FUNCTION F_EL6910MessageTemplate : STRING(255)
VAR_INPUT
    wTextId : WORD;
END_VAR

CASE wTextId OF
    16#0001: F_EL6910MessageTemplate := 'Primary MC: GLOBAL_Fault with Code 0x%x and Additional Code 0x%x';
    16#0002: F_EL6910MessageTemplate := 'Primary MC: GLOBAL_Shutdown with Code 0x%x and Additional Code 0x%x';
    16#0003: F_EL6910MessageTemplate := 'Secondary MC: GLOBAL_Fault with Code 0x%x and Additional Code 0x%x';
    16#0004: F_EL6910MessageTemplate := 'Secondary MC: GLOBAL_Shutdown with Code 0x%x and Additional Code 0x%x';
    16#0005: F_EL6910MessageTemplate := 'Primary MC: Stored GLOBAL_Fault with Code 0x%x and Additional Code 0x%x';
    16#0006: F_EL6910MessageTemplate := 'Secondary MC: Stored GLOBAL_Fault with Code 0x%x and Additional Code 0x%x';
    16#0007: F_EL6910MessageTemplate := 'Diag-Message-Overflow: %d messages got lost';
    16#0008: F_EL6910MessageTemplate := 'Primary MC: the CRC of the FRAM Data was wrong (Diag-Code=%d)';
    16#0009: F_EL6910MessageTemplate := 'Secondary MC: the CRC of the FRAM Data was wrong (Diag-Code=%d)';
    16#0010: F_EL6910MessageTemplate := 'Reserved CfgData has to be zero st offset %d';
    16#0011: F_EL6910MessageTemplate := 'The password is wrong';
    16#0012: F_EL6910MessageTemplate := 'The user was not found';
    16#0013: F_EL6910MessageTemplate := 'The CRC of the login data does not match';
    16#0014: F_EL6910MessageTemplate := 'The serial number of the login data does not match';
    16#0015: F_EL6910MessageTemplate := 'The login watchdog has been expired';
    16#0016: F_EL6910MessageTemplate := 'The user was logged out before';
    16#0017: F_EL6910MessageTemplate := 'The user has not sufficient access rights';
    16#0018: F_EL6910MessageTemplate := 'The reserved area of the CfgData was not 0';
    16#0019: F_EL6910MessageTemplate := 'The CRC of the CfgData was wrong';
    16#001A: F_EL6910MessageTemplate := 'The user name is wrong at word offset 0x%x when changing the password';
    16#001B: F_EL6910MessageTemplate := 'The requested number of users is too big';
    16#001D: F_EL6910MessageTemplate := 'The user update flags are wrong at word offset 0x%x when changing the password';
    16#001E: F_EL6910MessageTemplate := 'The wrong user (user %d) is logged in when changing the password (user %d found in the received data)';
    16#0021: F_EL6910MessageTemplate := 'the maximum Global-Shutdown counter was exceeded in the Vendor Data (maximum value: %d, actual value: %d)';
    16#0030: F_EL6910MessageTemplate := 'Sync Manager 2 Address (0x%x) is invalid, minimum value = 0x%x, maximum value = 0x%x';
    16#0031: F_EL6910MessageTemplate := 'Sync Manager 3 Address (0x%x) is invalid, minimum value = 0x%x, maximum value = 0x%x';
    16#0032: F_EL6910MessageTemplate := 'Sync Manager 4 Address (0x%x) is invalid, minimum value = 0x%x, maximum value = 0x%x';
    16#0033: F_EL6910MessageTemplate := 'Sync Manager 5 Address (0x%x) is invalid, minimum value = 0x%x, maximum value = 0x%x';
    16#0034: F_EL6910MessageTemplate := 'Sync Manager 2 Size (%d) is invalid, minimum value = %d, maximum value = %d';
    16#0035: F_EL6910MessageTemplate := 'Sync Manager 3 Size (%d) is invalid, minimum value = %d, maximum value = %d';
    16#0036: F_EL6910MessageTemplate := 'Sync Manager 4 Size (%d) is invalid, minimum value = %d, maximum value = %d';
    16#0037: F_EL6910MessageTemplate := 'Sync Manager 5 Size (%d) is invalid, minimum value = %d, maximum value = %d';
    16#0038: F_EL6910MessageTemplate := 'Sync Manager %d Settings (Offset 4-7) are invalid, expected values = 0x%x, 0x%x';
    16#0044: F_EL6910MessageTemplate := 'Sync Manager 6 Address (0x%x) is invalid, minimum value = 0x%x, maximum value = 0x%x';
    16#0045: F_EL6910MessageTemplate := 'Sync Manager 7 Address (0x%x) is invalid, minimum value = 0x%x, maximum value = 0x%x';
    16#0048: F_EL6910MessageTemplate := 'Sync Manager 6 Size (%d) is invalid, minimum value = %d, maximum value = %d';
    16#0049: F_EL6910MessageTemplate := 'Sync Manager 7 Size (%d) is invalid, minimum value = %d, maximum value = %d';
    16#0101: F_EL6910MessageTemplate := 'Primary MC: Completed RAM TEST: Starttime: 0x%x and Stoptime: 0x%x . The calculated timediff is 0x%x.';
    16#0102: F_EL6910MessageTemplate := 'Secondary MC: Completed RAM TEST: Starttime: 0x%x and Stoptime: 0x%x . The calculated timediff is 0x%x.';
    16#0115: F_EL6910MessageTemplate := 'Controller %d: Maximum temperature exceeded. Temperature is 0x%x, should be <= 0x%x.';
    16#0116: F_EL6910MessageTemplate := 'Controller %d: Minimum temperature alert. Temperature is 0x%x, should be >= 0x%x.';
    16#0117: F_EL6910MessageTemplate := 'Controller %d: Temperature difference too high. Difference is %d, should be <= %d.';
    16#0118: F_EL6910MessageTemplate := 'Controller %d: Maximum voltage alert (Partner_VCC). Voltage is 0x%x, should be <= 0x%x.';
    16#0119: F_EL6910MessageTemplate := 'Controller %d: Minimum voltage alert (Partner_VCC). Voltage is 0x%x, should be >= 0x%x.';
    16#011A: F_EL6910MessageTemplate := 'Controller %d: Maximum voltage alert (ECAT_VCC). Voltage is 0x%x, should be <= 0x%x.';
    16#011B: F_EL6910MessageTemplate := 'Controller %d: Minimum voltage alert (ECAT_VCC). Voltage is 0x%x, should be >= 0x%x.';
    16#011E: F_EL6910MessageTemplate := 'Controller %d: Timer Tick Difference is too high. Difference is 0x%x, should be >= 0x%x.';
    16#011F: F_EL6910MessageTemplate := 'Controller %d: Minimum value alert (Individual ADC Check). Channel parameter = %d. Actual value is 0x%x.';
    16#0120: F_EL6910MessageTemplate := 'Controller %d: Maximum value alert (Individual ADC Check). Channel parameter = %d. Actual value is 0x%x.';
    16#2001: F_EL6910MessageTemplate := 'The %d. connection has received an invalid FSoE-Cmd in state CONNECTION';
    16#2002: F_EL6910MessageTemplate := 'The %d. connection has received an unknown FSoE-Cmd in state CONNECTION';
    16#2003: F_EL6910MessageTemplate := 'The %d. connection has received an invalid FSoE-ConnID in state CONNECTION';
    16#2004: F_EL6910MessageTemplate := 'The %d. connection has received an invalid FSoE-CRC in state CONNECTION';
    16#2005: F_EL6910MessageTemplate := 'The FSoE-Watchdog of the %d. connection has been expired in state CONNECTION';
    16#2006: F_EL6910MessageTemplate := 'On the %d. connection the received FSoE-Address (0x%x) does not match with the expected FSoE-Address (0x%x)';
    16#2007: F_EL6910MessageTemplate := 'On the %d. connection the received connection data do not match with the sent values';
    16#200C: F_EL6910MessageTemplate := 'On the %d. connection in state CONNECTION the Connection was restarted from the FSoE-Master';
    16#200E: F_EL6910MessageTemplate := 'A Module fault was detected on the %d. connection in state CONNECTION';
    16#2011: F_EL6910MessageTemplate := 'On the %d. connection in state CONNECTION a FSoE-Reset with Error-Code 1 was received which means that the communication partner has received an invalid FSoE-Cmd';
    16#2012: F_EL6910MessageTemplate := 'On the %d. connection in state CONNECTION a FSoE-Reset with Error-Code 2 was received which means that the communication partner has received an unknown FSoE-Cmd';
    16#2013: F_EL6910MessageTemplate := 'On the %d. connection in state CONNECTION a FSoE-Reset with Error-Code 3 was received which means that the communication partner has received an invalid FSoE-ConnID';
    16#2014: F_EL6910MessageTemplate := 'On the %d. connection in state CONNECTION a FSoE-Reset with Error-Code 4 was received which means that the communication partner has received an invalid FSoE-CRC';
    16#2015: F_EL6910MessageTemplate := 'On the %d. connection in state CONNECTION a FSoE-Reset with Error-Code 5 was received which means that the FSoE-Watchdog has been expired in the communication partner';
    16#2016: F_EL6910MessageTemplate := 'On the %d. connection in state CONNECTION a FSoE-Reset with Error-Code 6 was received which means that the communication partner has received an invalid FSoE-Address';
    16#2017: F_EL6910MessageTemplate := 'On the %d. connection in state CONNECTION a FSoE-Reset with Error-Code 7 was received which means that the communication partner has received connection data do not match with the sent values';
    16#2018: F_EL6910MessageTemplate := 'On the %d. connection in state CONNECTION a FSoE-Reset with Error-Code 8 was received which means that the communication partner has received an invalid communication parameter length';
    16#2019: F_EL6910MessageTemplate := 'On the %d. connection in state CONNECTION a FSoE-Reset with Error-Code 9 was received which means that the communication partner has received an invalid FSoE Watchdog';
    16#201A: F_EL6910MessageTemplate := 'On the %d. connection in state CONNECTION a FSoE-Reset with Error-Code 10 was received which means that the communication partner has received an invalid application parameter length';
    16#201B: F_EL6910MessageTemplate := 'On the %d. connection in state CONNECTION a FSoE-Reset with Error-Code 11 was received which means that the communication partner has received invalid application parameter data';
    16#201C: F_EL6910MessageTemplate := 'On the %d. connection in state CONNECTION a FSoE-Reset with Error-Code 12 was received';
    16#201D: F_EL6910MessageTemplate := 'On the %d. connection in state CONNECTION a FSoE-Reset with Error-Code 13 was received';
    16#201E: F_EL6910MessageTemplate := 'On the %d. connection in state CONNECTION a FSoE-Reset with Error-Code 14 was received which means that the communication partner has detected a module fault';
    16#201F: F_EL6910MessageTemplate := 'On the %d. connection in state CONNECTION a FSoE-Reset with Error-Code 0x%x was received';
    16#2041: F_EL6910MessageTemplate := 'The %d. connection has received an invalid FSoE-Cmd in state PARAMETER';
    16#2042: F_EL6910MessageTemplate := 'The %d. connection has received an unknown FSoE-Cmd in state PARAMETER';
    16#2043: F_EL6910MessageTemplate := 'The %d. connection has received an invalid FSoE-ConnID in state PARAMETER';
    16#2044: F_EL6910MessageTemplate := 'The %d. connection has received an invalid FSoE-CRC in state PARAMETER';
    16#2045: F_EL6910MessageTemplate := 'The FSoE-Watchdog of the %d. connection has been expired in state PARAMETER';
    16#2047: F_EL6910MessageTemplate := 'On the %d. connection the received parameter data do not match with the sent values';
    16#2048: F_EL6910MessageTemplate := 'On the %d. connection the received communication parameter length (%d) does not match with the expected value of 2';
    16#2049: F_EL6910MessageTemplate := 'On the %d. connection the received FSoE Watchdog (%d) is outside the allowed area from 2 to 60000';
    16#204A: F_EL6910MessageTemplate := 'On the %d. connection the received application parameter length (%d) is unequal the expected length of %d';
    16#204B: F_EL6910MessageTemplate := 'On the %d. connection the received application parameter data are wrong';
    16#204C: F_EL6910MessageTemplate := 'On the %d. connection in state PARAMETER the Connection was restarted from the FSoE-Master';
    16#204E: F_EL6910MessageTemplate := 'A Module fault was detected on the %d. connection in state PARAMETER';
    16#2051: F_EL6910MessageTemplate := 'On the %d. connection in state PARAMETER a FSoE-Reset with Error-Code 1 was received which means that the communication partner has received an invalid FSoE-Cmd';
    16#2052: F_EL6910MessageTemplate := 'On the %d. connection in state PARAMETER a FSoE-Reset with Error-Code 2 was received which means that the communication partner has received an unknown FSoE-Cmd';
    16#2053: F_EL6910MessageTemplate := 'On the %d. connection in state PARAMETER a FSoE-Reset with Error-Code 3 was received which means that the communication partner has received an invalid FSoE-ConnID';
    16#2054: F_EL6910MessageTemplate := 'On the %d. connection in state PARAMETER a FSoE-Reset with Error-Code 4 was received which means that the communication partner has received an invalid FSoE-CRC';
    16#2055: F_EL6910MessageTemplate := 'On the %d. connection in state PARAMETER a FSoE-Reset with Error-Code 5 was received which means that the FSoE-Watchdog has been expired in the communication partner';
    16#2056: F_EL6910MessageTemplate := 'On the %d. connection in state PARAMETER a FSoE-Reset with Error-Code 6 was received which means that the communication partner has received an invalid FSoE-Address';
    16#2057: F_EL6910MessageTemplate := 'On the %d. connection in state PARAMETER a FSoE-Reset with Error-Code 7 was received which means that the communication partner has received connection data do not match with the sent values';
    16#2058: F_EL6910MessageTemplate := 'On the %d. connection in state PARAMETER a FSoE-Reset with Error-Code 8 was received which means that the communication partner has received an invalid communication parameter length';
    16#2059: F_EL6910MessageTemplate := 'On the %d. connection in state PARAMETER a FSoE-Reset with Error-Code 9 was received which means that the communication partner has received an invalid FSoE Watchdog';
    16#205A: F_EL6910MessageTemplate := 'On the %d. connection in state PARAMETER a FSoE-Reset with Error-Code 10 was received which means that the communication partner has received an invalid application parameter length';
    16#205B: F_EL6910MessageTemplate := 'On the %d. connection in state PARAMETER a FSoE-Reset with Error-Code 11 was received which means that the communication partner has received invalid application parameter data';
    16#205C: F_EL6910MessageTemplate := 'On the %d. connection in state PARAMETER a FSoE-Reset with Error-Code 12 was received';
    16#205D: F_EL6910MessageTemplate := 'On the %d. connection in state PARAMETER a FSoE-Reset with Error-Code 13 was received';
    16#205E: F_EL6910MessageTemplate := 'On the %d. connection in state PARAMETER a FSoE-Reset with Error-Code 14 was received which means that the communication partner has detected a module fault';
    16#205F: F_EL6910MessageTemplate := 'On the %d. connection in state PARAMETER a FSoE-Reset with Error-Code 0x%x was received';
    16#2061: F_EL6910MessageTemplate := 'On the %d. connection in state PARAMETER a wrong Command was received, which means that the Safe-Parameter size is wrong (Expected size: %d, Received size: %d)';
    16#2081: F_EL6910MessageTemplate := 'The %d. connection has received an invalid FSoE-Cmd in state DATA';
    16#2082: F_EL6910MessageTemplate := 'The %d. connection has received an unknown FSoE-Cmd in state DATA';
    16#2083: F_EL6910MessageTemplate := 'The %d. connection has received an invalid FSoE-ConnID in state DATA';
    16#2084: F_EL6910MessageTemplate := 'The %d. connection has received an invalid FSoE-CRC in state DATA';
    16#2085: F_EL6910MessageTemplate := 'The FSoE-Watchdog of the %d. connection has been expired in state DATA';
    16#208C: F_EL6910MessageTemplate := 'On the %d. connection in state DATA the Connection was restarted from the FSoE-Master';
    16#208D: F_EL6910MessageTemplate := 'The FailSafeData command was received on the %d. connection in state DATA';
    16#208E: F_EL6910MessageTemplate := 'A Module fault was detected on the %d. connection in state DATA';
    16#2091: F_EL6910MessageTemplate := 'On the %d. connection in state DATA a FSoE-Reset with Error-Code 1 was received which means that the communication partner has received an invalid FSoE-Cmd';
    16#2092: F_EL6910MessageTemplate := 'On the %d. connection in state DATA a FSoE-Reset with Error-Code 2 was received which means that the communication partner has received an unknown FSoE-Cmd';
    16#2093: F_EL6910MessageTemplate := 'On the %d. connection in state DATA a FSoE-Reset with Error-Code 3 was received which means that the communication partner has received an invalid FSoE-ConnID';
    16#2094: F_EL6910MessageTemplate := 'On the %d. connection in state DATA a FSoE-Reset with Error-Code 4 was received which means that the communication partner has received an invalid FSoE-CRC';
    16#2095: F_EL6910MessageTemplate := 'On the %d. connection in state DATA a FSoE-Reset with Error-Code 5 was received which means that the FSoE-Watchdog has been expired in the communication partner';
    16#2096: F_EL6910MessageTemplate := 'On the %d. connection in state DATA a FSoE-Reset with Error-Code 6 was received which means that the communication partner has received an invalid FSoE-Address';
    16#2097: F_EL6910MessageTemplate := 'On the %d. connection in state DATA a FSoE-Reset with Error-Code 7 was received which means that the communication partner has received connection data do not match with the sent values';
    16#2098: F_EL6910MessageTemplate := 'On the %d. connection in state DATA a FSoE-Reset with Error-Code 8 was received which means that the communication partner has received an invalid communication parameter length';
    16#2099: F_EL6910MessageTemplate := 'On the %d. connection in state DATA a FSoE-Reset with Error-Code 9 was received which means that the communication partner has received an invalid FSoE Watchdog';
    16#209A: F_EL6910MessageTemplate := 'On the %d. connection in state DATA a FSoE-Reset with Error-Code 10 was received which means that the communication partner has received an invalid application parameter length';
    16#209B: F_EL6910MessageTemplate := 'On the %d. connection in state DATA a FSoE-Reset with Error-Code 11 was received which means that the communication partner has received invalid application parameter data';
    16#209C: F_EL6910MessageTemplate := 'On the %d. connection in state DATA a FSoE-Reset with Error-Code 12 was received';
    16#209D: F_EL6910MessageTemplate := 'On the %d. connection in state DATA a FSoE-Reset with Error-Code 13 was received';
    16#209E: F_EL6910MessageTemplate := 'On the %d. connection in state DATA a FSoE-Reset with Error-Code 14 was received which means that the communication partner has detected a module fault';
    16#209F: F_EL6910MessageTemplate := 'On the %d. connection in state DATA a FSoE-Reset with Error-Code 0x%x was received';
    16#20C1: F_EL6910MessageTemplate := 'The %d. connection has received an invalid FSoE-Cmd in state SHUTDOWN';
    16#20C2: F_EL6910MessageTemplate := 'The %d. connection has received an unknown FSoE-Cmd in state SHUTDOWN';
    16#20C4: F_EL6910MessageTemplate := 'The %d. connection has received an invalid FSoE-CRC in state SHUTDOWN';
    16#20E3: F_EL6910MessageTemplate := 'The %d. connection has received the invalid FSoE-ConnID 0 in state SESSION';
    16#2101: F_EL6910MessageTemplate := 'On the %d. connection the PROFIsafe-Slave reports a communication error';
    16#2102: F_EL6910MessageTemplate := 'On the %d. connection the PROFIsafe-Slave reports a watchdog error';
    16#2103: F_EL6910MessageTemplate := 'On the %d. connection the PROFIsafe-Slave reports a device fault';
    16#2104: F_EL6910MessageTemplate := 'On the %d. connection a CRC2-Error was detected locally on the PROFIsafe Host';
    16#2105: F_EL6910MessageTemplate := 'On the %d. connection the Watchdog has been expired locally on the PROFIsafe Host';
    16#2114: F_EL6910MessageTemplate := 'On the %d. connection a CRC2-Error was detected locally on the PROFIsafe Slave';
    16#2115: F_EL6910MessageTemplate := 'On the %d. connection the Watchdog has been expired locally on the PROFIsafe Slave';
    16#2117: F_EL6910MessageTemplate := 'On the %d. connection the Bit 7 of the F_Control is reset, which is not allowed on a PROFIsafe Slave connection with the same message size for inputs and outputs';
    16#211C: F_EL6910MessageTemplate := 'On the %d. connection the PROFIsafe Slave has been restarted locally';
    16#3000: F_EL6910MessageTemplate := 'The received number of groups (%d) was too big, the maximum allowed value is %d';
    16#3001: F_EL6910MessageTemplate := 'The received number of FBs (%d) was too big, the maximum allowed value is %d';
    16#3002: F_EL6910MessageTemplate := 'The received number of Connections (%d) was too big, the maximum allowed value is %d';
    16#3003: F_EL6910MessageTemplate := 'The received number of Output Mappings was too big, the maximum allowed value is %d';
    16#3004: F_EL6910MessageTemplate := 'The received number of Input Mappings was too big, the maximum allowed value is %d';
    16#3005: F_EL6910MessageTemplate := 'The received size of Standard Inputs (%d) was too big, the maximum allowed value is %d';
    16#3006: F_EL6910MessageTemplate := 'The received size of Standard Outputs (%d) was too big, the maximum allowed value is %d';
    16#3007: F_EL6910MessageTemplate := 'The received number of Restore Slaves (%d) was too big, the maximum allowed value is %d';
    16#3008: F_EL6910MessageTemplate := 'The SafeCfgData type was unexpected: %d found and %d expected';
    16#3009: F_EL6910MessageTemplate := 'The SafeCfgData type 2 (Connection) was expected at offset %d';
    16#300A: F_EL6910MessageTemplate := 'The SafeCfgData type 3 (FB) was expected at offset %d';
    16#300B: F_EL6910MessageTemplate := 'The SafeCfgData type 15 (GAP) was expected at offset %d';
    16#300C: F_EL6910MessageTemplate := 'The Bit-Mask in the SafeCfgData was wrong at offset %d';
    16#300D: F_EL6910MessageTemplate := 'The address in the SafeCfgData was wrong at offset %d';
    16#300E: F_EL6910MessageTemplate := 'The Signal number in the SafeCfgData was wrong at offset %d';
    16#300F: F_EL6910MessageTemplate := 'The number of connections was wrong in the SafeCfgData of the Group at offset %d';
    16#3010: F_EL6910MessageTemplate := 'The number of FBs was wrong in the SafeCfgData of the Group at offset %d';
    16#3011: F_EL6910MessageTemplate := 'The size of the SafeCfgData was wrong at offset %d';
    16#3012: F_EL6910MessageTemplate := 'The complete size of the SafeCfgData related to the Group %d was wrong';
    16#3013: F_EL6910MessageTemplate := 'If the RUN-Signal should be mapped internally, it has to be activated at offset %d';
    16#3014: F_EL6910MessageTemplate := 'The message size at offset %d is invalid';
    16#3015: F_EL6910MessageTemplate := 'The connection parameter at offset %d is invalid';
    16#3016: F_EL6910MessageTemplate := 'If the ERRACK-Signal should be mapped internally, it has to be activated at offset %d';
    16#3017: F_EL6910MessageTemplate := 'The connection type at offset %d is invalid';
    16#3018: F_EL6910MessageTemplate := 'The value at offset %d of the SafeCfgData is invalid';
    16#3019: F_EL6910MessageTemplate := 'The value at offset %d of the SafeCfgData is invalid because at least one of the related signals is not active';
    16#301A: F_EL6910MessageTemplate := 'The number of mappings (%d) is wrong because it is not the last Mapping SafeCfgData';
    16#301B: F_EL6910MessageTemplate := 'The Safe Logic Cfg Data were downloaded in the wrong download state (%d)';
    16#301C: F_EL6910MessageTemplate := 'The number of mappings (%d) is too great in the Mapping SafeCfgData';
    16#301D: F_EL6910MessageTemplate := 'The Mapping-Size in the SafeCfgData was wrong at offset %d';
    16#301E: F_EL6910MessageTemplate := 'A Group-Input Mapping was expected at offset %d';
    16#301F: F_EL6910MessageTemplate := 'A Connection-Input Mapping was expected at offset %d';
    16#3020: F_EL6910MessageTemplate := 'A FB-Input Bit-Mapping was expected at offset %d';
    16#3021: F_EL6910MessageTemplate := 'A FB-Input Byte-Mapping was expected at offset %d';
    16#3022: F_EL6910MessageTemplate := 'No more mapping was expected at offset %d';
    16#3023: F_EL6910MessageTemplate := 'Invalid Safe User Parameter size at byte offset 0x%x (Found=%d, Expected=%d)';
    16#3024: F_EL6910MessageTemplate := 'The SafeCfgData type 4 (Safe User Parameter) was expected at offset %d';
    16#3025: F_EL6910MessageTemplate := 'The download of the Input Mapping Cfg Data was refused because %d groups were missing in the Safe Logic Cfg Data';
    16#3026: F_EL6910MessageTemplate := 'The download of the Input Mapping Cfg Data was refused because %d connections were missing in the Safe Logic Cfg Data';
    16#3027: F_EL6910MessageTemplate := 'The download of the Input Mapping Cfg Data was refused because %d FBs were missing in the Safe Logic Cfg Data';
    16#3028: F_EL6910MessageTemplate := 'At least one group has to be defined in the SafeCfgData';
    16#3029: F_EL6910MessageTemplate := 'The download of the Input Mapping Cfg Data was refused because no safe Logic Cfg Data were downloaded before';
    16#302A: F_EL6910MessageTemplate := 'The Subindex %d was expected to be downloaded';
    16#302B: F_EL6910MessageTemplate := 'When loading CfgData a user has to be logged in before';
    16#302C: F_EL6910MessageTemplate := 'The Input Mapping Cfg Data were downloaded in the wrong download state (%d)';
    16#302D: F_EL6910MessageTemplate := 'The download of theSafe Logic CfgData is refused because the old Safe Logic Cfg Data were not deleted before';
    16#302E: F_EL6910MessageTemplate := 'The user was logged out before';
    16#302F: F_EL6910MessageTemplate := 'The user has not sufficient access rights';
    16#3030: F_EL6910MessageTemplate := 'The reserved area of the CfgData was not 0';
    16#3031: F_EL6910MessageTemplate := 'The CRC of the CfgData was wrong';
    16#3032: F_EL6910MessageTemplate := 'All needed CfgData pages were downloaded before, no more pages are expected';
    16#3033: F_EL6910MessageTemplate := 'The mapping code buffer is too small for the mapping (Offset: 0x%x, Size: %d)';
    16#3034: F_EL6910MessageTemplate := 'The maximum allowed subindex is %d';
    16#3035: F_EL6910MessageTemplate := 'The download of the Output Mapping Cfg Data was refused because %d mappings of the Input Mapping Cfg Data were missing';
    16#3036: F_EL6910MessageTemplate := '%d input mappings of the groups were missing in the Input Mapping Cfg Data';
    16#3037: F_EL6910MessageTemplate := '%d input mappings of the connections were missing in the Input Mapping Cfg Data';
    16#3038: F_EL6910MessageTemplate := '%d input bit mappings of the FBs were missing in the Input Mapping Cfg Data';
    16#3039: F_EL6910MessageTemplate := '%d input byte mappings of the FBs were missing in the Input Mapping Cfg Data';
    16#303A: F_EL6910MessageTemplate := 'The Output Mapping Cfg Data were downloaded in the wrong download state (%d)';
    16#303B: F_EL6910MessageTemplate := 'The mapping code buffer is too small for the local mapping';
    16#303C: F_EL6910MessageTemplate := 'The download of the Safe Parameter was refused because no Output Mapping Cfg Data were downloaded before';
    16#303D: F_EL6910MessageTemplate := 'The download of the Safe User Parameter was refused because %d mappings of the Output Mapping Cfg Data were missing';
    16#303E: F_EL6910MessageTemplate := 'The Safe User Parameter Cfg Data were downloaded in the wrong download state (%d)';
    16#303F: F_EL6910MessageTemplate := 'The download of the Activate Project Cfg Data was refused because no Safe User Parameter Cfg Data were downloaded before';
    16#3040: F_EL6910MessageTemplate := 'The download of the Activate Project Cfg Data was refused because %d bytes of the Safe Parameter Cfg Data were missing';
    16#3041: F_EL6910MessageTemplate := 'The received activate code (0x%x) was wrong in the Project Cfg Data';
    16#3042: F_EL6910MessageTemplate := 'The TwinSAFE Address (%d) in the Project Cfg Data does not match with the DIP switch (%d)';
    16#3043: F_EL6910MessageTemplate := 'At least one Cfg Data page has to be defined in the Safe Logic Cfg Data';
    16#3044: F_EL6910MessageTemplate := 'The maximum number (%d) of Cfg Data pages was exceeded in the Safe Logic Cfg Data';
    16#3045: F_EL6910MessageTemplate := 'The received number of Safe Logic Cfg Data pages (%d) has exceeded the configured value at offset 0 of the Safe Logic Cfg Data (%d)';
    16#3046: F_EL6910MessageTemplate := 'The download of the Input Mapping Cfg Data was refused because %d pages were missing in the Safe Logic Cfg Data';
    16#3047: F_EL6910MessageTemplate := 'The Safe Logic Cfg Data CRC does not match in the Safe Project Cfg Data';
    16#3048: F_EL6910MessageTemplate := 'When checking the Mapping Code a fault has detected at offset 0x%x';
    16#3049: F_EL6910MessageTemplate := 'The Mapping Cfg Data CRC does not match in the Safe Project Cfg Data';
    16#304A: F_EL6910MessageTemplate := 'The number of Input Mappings is too small in the Safe Project Cfg Data (Code-Offset=0x%x)';
    16#304B: F_EL6910MessageTemplate := 'The number of Output Mappings is too small in the Safe Project Cfg Data (Code-Offset=0x%x)';
    16#304C: F_EL6910MessageTemplate := 'The number of Input Mappings is too great in the Safe Project Cfg Data, (%d mappings too much, Code-Offset=0x%x)';
    16#304D: F_EL6910MessageTemplate := 'The number of Output Mappings is too great in the Safe Project Cfg Data, (%d mappings too much, Code-Offset=0x%x)';
    16#304E: F_EL6910MessageTemplate := 'The maximum number (%d) of Cfg Data pages was exceeded in the Safe User Parameter Cfg Data';
    16#304F: F_EL6910MessageTemplate := 'At least one Cfg Data page has to be defined in the Safe User Parameter Cfg Data';
    16#3050: F_EL6910MessageTemplate := 'The Safe User Parameter Cfg Data CRC does not match in the Safe Project Cfg Data';
    16#3052: F_EL6910MessageTemplate := 'The calculated local process image size (%d) exceeded the maximum local process image size of %d';
    16#3053: F_EL6910MessageTemplate := 'The Activate Project Cfg Data were downloaded in the wrong download state (%d)';
    16#3054: F_EL6910MessageTemplate := 'The Delete Project Cfg Data were downloaded in the wrong download state (%d)';
    16#3055: F_EL6910MessageTemplate := 'The TwinSAFE Address (%d) does not match with the DIP switch (%d) in the Delete Project Cfg Data';
    16#3056: F_EL6910MessageTemplate := 'The Delete Code (%d) is too high in the Delete Project Cfg Data';
    16#3057: F_EL6910MessageTemplate := 'Unexpected connection index in the Safe User Parameter Cfg Data at byte offset 0x%x';
    16#3058: F_EL6910MessageTemplate := 'The received number of Local Safety Inputs (%d) was wrong, the expected value is %d';
    16#3059: F_EL6910MessageTemplate := 'The received number of Local Safety Outputs (%d) was wrong, the expected value is %d';
    16#305A: F_EL6910MessageTemplate := 'The received number of Local Standard Inputs (%d) was wrong, the expected value is %d';
    16#305B: F_EL6910MessageTemplate := 'The received number of Local Standard Outputs (%d) was wrong, the expected value is %d';
    16#305C: F_EL6910MessageTemplate := 'The received Safety Input Message size at word offset 15 of the Safe Logic Cfg Data (%d) is unequal the calculated value of %d';
    16#305D: F_EL6910MessageTemplate := 'The received Safety Output Message size at word offset 16 of the Safe Logic Cfg Data (%d) is unequal the calculated value of %d';
    16#305E: F_EL6910MessageTemplate := 'The received Safety Input size at word offset 7 of the Safe Logic Cfg Data (%d) is unequal the calculated value of %d';
    16#305F: F_EL6910MessageTemplate := 'The received Safety Output size at word offset 8 of the Safe Logic Cfg Data (%d) is unequal the calculated value of %d';
    16#3060: F_EL6910MessageTemplate := 'The received PROFIsafe Input Message size at word offset 9 of the Safe Logic Cfg Data (%d) is unequal the calculated value of %d';
    16#3061: F_EL6910MessageTemplate := 'The received PROFIsafe Output Message size at word offset 10 of the Safe Logic Cfg Data (%d) is unequal the calculated value of %d';
    16#3062: F_EL6910MessageTemplate := 'At word offset 0x%x the configured number of CRCs of %d exceeds the maximum number of CRCs (%d)';
    16#3063: F_EL6910MessageTemplate := 'The received SafeUserParameterSizeInFrame (%d) was wrong, the expected value is %d';
    16#3064: F_EL6910MessageTemplate := 'The received FB Analog Input size at word offset 13 of the Safe Logic Cfg Data (%d) is unequal the calculated value of %d';
    16#3065: F_EL6910MessageTemplate := 'The received FB Analog Output size at word offset 14 of the Safe Logic Cfg Data (%d) is unequal the calculated value of %d';
    16#3066: F_EL6910MessageTemplate := 'The received Connection Status Data size at word offset 21 of the Safe Logic Cfg Data (%d) is unequal the calculated value of %d';
    16#3067: F_EL6910MessageTemplate := 'The received FB Status Data size at word offset 22 of the Safe Logic Cfg Data (%d) is unequal the calculated value of %d';
    16#3068: F_EL6910MessageTemplate := 'The number of active signals in the FB is invalid at offset %d';
    16#3069: F_EL6910MessageTemplate := 'The local map code size in the FB is invalid at offset %d';
    16#306A: F_EL6910MessageTemplate := 'The analog output size in the Group Cfg Data is invalid at offset %d';
    16#306B: F_EL6910MessageTemplate := 'The analog output offset in the Group Cfg Data is invalid at offset %d';
    16#306C: F_EL6910MessageTemplate := 'The received FB Analog Output size at word offset 14 of the Safe Logic Cfg Data (%d) is unequal the calculated value over all the Group Cfg Data (%d)';
    16#306D: F_EL6910MessageTemplate := 'The calculated end of the analog output area (%d) is unequal the calculated analog output offset over all the Group Cfg Data (%d)';
    16#306E: F_EL6910MessageTemplate := 'The value of the FB Cfg Data at offset %d is invalid';
    16#306F: F_EL6910MessageTemplate := 'At least one FB input has to be deactivated in this operation mode at offset %d';
    16#3070: F_EL6910MessageTemplate := 'At least the level of one FB input is wrong in this operation mode at offset %d';
    16#3071: F_EL6910MessageTemplate := 'The value of the FB Cfg Data at word offset %d is invalid in this operation mode';
    16#3072: F_EL6910MessageTemplate := 'The number (%d) of Cfg Data pages was exceeded in the Info Data Cfg Data at offset 0';
    16#3073: F_EL6910MessageTemplate := 'The received number of FBs (%d) at word offset 1 was unequal the configured number of FBs of %d';
    16#3074: F_EL6910MessageTemplate := 'The received FB Status Data Size (%d) in the Info Data Map Cfg Data at byte offset %d is unequal the calculated FB Status Data size of %d';
    16#3075: F_EL6910MessageTemplate := 'The received FB Diag Data Size (%d) in the Info Data Map Cfg Data at byte offset %d is unequal the calculated FB Diag Data size of %d';
    16#3076: F_EL6910MessageTemplate := 'The received number of Connections (%d) in the Info Data Cfg Data at word offset %d was unequal the configured number of connections of %d';
    16#3077: F_EL6910MessageTemplate := 'The received Connection Type (%d) in the Info Data Map Cfg Data at byte offset %d is unequal the configured Connection Type of %d';
    16#3078: F_EL6910MessageTemplate := 'The FB Diag Data Map in the Info Data Map Cfg Data was wrong at byte offset %d (bit 7=1 and bit 6=0 is not allowed)';
    16#3079: F_EL6910MessageTemplate := 'The received number of Groups (%d) in the Info Data Cfg Data at word offset %d was unequal the configured number of Groups of %d';
    16#307A: F_EL6910MessageTemplate := 'The FB-Type is unknown at offset 0x%x';
    16#307B: F_EL6910MessageTemplate := 'The value at offset %d of the SafeCfgData is too great';
    16#307C: F_EL6910MessageTemplate := 'The value at offset %d of the SafeCfgData is too small';
    16#307D: F_EL6910MessageTemplate := 'FB-Muting: if SequentialInputs is TRUE, all MuteIn signals have to be active at offset 0x%x';
    16#307E: F_EL6910MessageTemplate := 'The type of the analog inputs has to be the same at offset 0x%x';
    16#307F: F_EL6910MessageTemplate := 'The received size of the local safe user parameter (%d) was wrong, the expected size is %d';
    16#3080: F_EL6910MessageTemplate := 'The value at offset %d of the SafeCfgData is invalid in combination with the value %d words before in the SafeCfgData';
    16#3081: F_EL6910MessageTemplate := 'The received size of the FB Parameter Data at word offset 25 of the Safe Logic Cfg Data (%d) is unequal the calculated value of %d';
    16#3082: F_EL6910MessageTemplate := 'The FB-Type in the Change FB Parameter Data (FB %d) is unequal, the expected FB-type is %d';
    16#3083: F_EL6910MessageTemplate := 'The size in the Change FB Parameter Data (FB %d) is unequal, the expected size is %d';
    16#3084: F_EL6910MessageTemplate := 'The Setting Mode of the FB CAMMON (FB %d) in the Change FB Parameter Data is not activated';
    16#3085: F_EL6910MessageTemplate := 'The actual Logic State (%d) is unequal RUN (1) when changing FB Parameter Data';
    16#3086: F_EL6910MessageTemplate := 'The FB-Number (%d) in the Change FB Parameter Data is invalid';
    16#3087: F_EL6910MessageTemplate := 'The FRAM data size (%d) has exceeded, the maximum allowed value is %d';
    16#3088: F_EL6910MessageTemplate := 'The Safe User Parameter in the Change FB Parameter Data are not supported';
    16#3089: F_EL6910MessageTemplate := 'The size (%d) of the Change FB Parameter Data is too small, %d bytes are expected';
    16#308A: F_EL6910MessageTemplate := 'The type (%d) of the Safe User Parameter in the Change FB Parameter Data is wrong';
    16#308B: F_EL6910MessageTemplate := 'The size (%d) of the Safe User Parameter in the Change FB Parameter Data is wrong, the expected size is %d';
    16#308C: F_EL6910MessageTemplate := 'The offset of the Cyclic FRAM Data was wrong at offset %d';
    16#308D: F_EL6910MessageTemplate := 'No Local Input bytes configured for Extended Info Data Mapping';
    16#308E: F_EL6910MessageTemplate := 'No Local Output bytes configured for Extended Info Data Mapping';
    16#308F: F_EL6910MessageTemplate := 'Too much Local Input bytes configured for Info Data, only 31 bytes are allowed';
    16#3090: F_EL6910MessageTemplate := 'Too much Local Output bytes configured for Info Data, only 31 bytes are allowed';
    16#3094: F_EL6910MessageTemplate := 'The size 0 is not allowed for the safe user parameter at word offset %d';
    16#3095: F_EL6910MessageTemplate := 'The download of the Activate Project Cfg Data was refused because no Output Mapping Cfg Data were downloaded before';
    16#3096: F_EL6910MessageTemplate := 'The download of the Activate Project Cfg Data was refused because %d mappings of the Output Mapping Cfg Data were missing';
    16#3097: F_EL6910MessageTemplate := 'The re-converted FB-Mapping-Code was not matching to the FB Cfg Data (FB: %d, Code-Address: 0x%x, Offset: 0x%x)';
    16#3098: F_EL6910MessageTemplate := 'a destination was mapped twice in the bit mapping code (page: 0x%x, Code-Address: 0x%x)';
    16#3099: F_EL6910MessageTemplate := 'a destination was mapped twice in the byte mapping code (Page: 0x%x, Code-Address: 0x%x)';
    16#309A: F_EL6910MessageTemplate := 'the number of groups was exceeded in the Vendor Data (actual value: %d, minimum: %d, maximum: %d)';
    16#309B: F_EL6910MessageTemplate := 'the number of FBs was exceeded in the Vendor Data (actual value: %d, minimum: %d, maximum: %d)';
    16#309C: F_EL6910MessageTemplate := 'the number of Connections was exceeded in the Vendor Data (actual value: %d, minimum: %d, maximum: %d)';
    16#309D: F_EL6910MessageTemplate := 'the number of Standard Inputs was exceeded in the Vendor Data (actual value: %d, minimum: %d, maximum: %d)';
    16#309E: F_EL6910MessageTemplate := 'the number of Standard Outputs was exceeded in the Vendor Data (actual value: %d, minimum: %d, maximum: %d)';
    16#309F: F_EL6910MessageTemplate := 'the FSoE message size was exceeded in the Vendor Data (actual value: %d, minimum: %d, maximum: %d)';
    16#30A0: F_EL6910MessageTemplate := 'the FSoE safe user parameter size was exceeded in the Vendor Data (actual value: %d, minimum: %d, maximum: %d)';
    16#30A1: F_EL6910MessageTemplate := 'the PROFIsafe message size was exceeded in the Vendor Data (actual value: %d, minimum: %d, maximum: %d)';
    16#30A2: F_EL6910MessageTemplate := 'the EtherCAT Output size was exceeded in the Vendor Data (actual value: %d, minimum: %d, maximum: %d)';
    16#30A3: F_EL6910MessageTemplate := 'the EtherCAT Input size was exceeded in the Vendor Data (actual value: %d, minimum: %d, maximum: %d)';
    16#30A4: F_EL6910MessageTemplate := 'the EtherCAT Output size was exceeded in the project (calculated value: %d, maximum value: %d)';
    16#30A5: F_EL6910MessageTemplate := 'the EtherCAT Input size was exceeded in the project (calculated value: %d, maximum value: %d)';
    16#30A6: F_EL6910MessageTemplate := 'when re-converting the local FB mapping code (FB %d) the analog destination address was below the minimum value (Code-Offset: 0x%x, Data-Offset: 0x%x)';
    16#30A7: F_EL6910MessageTemplate := 'when re-converting the local FB mapping code (FB %d) the analog destination address was above the maximum value (Code-Offset: 0x%x, Data-Offset: 0x%x)';
    16#30A8: F_EL6910MessageTemplate := 'when re-converting the local FB mapping code (FB %d) the destination address was not found (Code-Offset: 0x%x, Data-Offset: 0x%x)';
    16#30A9: F_EL6910MessageTemplate := 'when re-converting the local FB mapping code (FB %d) the digital destination address was below the minimum value (Code-Offset: 0x%x, Data-Offset: 0x%x)';
    16#30AA: F_EL6910MessageTemplate := 'when re-converting the local FB mapping code (FB %d) the digital destination address was above the maximum value (Code-Offset: 0x%x, Data-Offset: 0x%x)';
    16#30AB: F_EL6910MessageTemplate := 'when re-converting the local FB mapping code (FB %d) the generated mapping data size was wrong (Code-Offset: 0x%x)';
    16#30AC: F_EL6910MessageTemplate := 'the Project CRC in the Activate Project Cfg Data was wrong';
    16#30AD: F_EL6910MessageTemplate := 'when re-converting the local FB mapping code the source bit address was wrong (FB: %d, Code-Offset: 0x%x)';
    16#30AE: F_EL6910MessageTemplate := 'when re-converting the local FB mapping code the source byte address was wrong (FB: %d, Code-Offset: 0x%x)';
    16#30B1: F_EL6910MessageTemplate := 'wrong subindex order when reading the input mapping cfg data, the expected subindex is %d';
    16#30B2: F_EL6910MessageTemplate := 'subindex exceeded when reading the cfg data';
    16#30B3: F_EL6910MessageTemplate := 'the offset in the Replacement Values cfg data is wrong in the Group cfg data at word-offset 0x%x';
    16#30B4: F_EL6910MessageTemplate := 'the deactivation mode passivate is enabled and the number of connections is unequal 1 in the Group cfg data at word-offset 0x%x';
    16#30B5: F_EL6910MessageTemplate := 'the RUN-signal has to be active in the Group cfg data at word-offset 0x%x';
    16#30B6: F_EL6910MessageTemplate := 'in the Change FB-Parameter (FB %d) the FB-type %d is not supported';
    16#30B7: F_EL6910MessageTemplate := 'the Subindex exceeds the number of connections (%d) when writing the PROFIsafe F-Parameter';
    16#30B8: F_EL6910MessageTemplate := 'the Connection-Type %d does not support PROFIsafe F-Parameter';
    16#30B9: F_EL6910MessageTemplate := 'the Subindex exceeds the number of connections (%d) when writing the Store Slave Project CRC Parameter';
    16#30BA: F_EL6910MessageTemplate := 'the Connection-Type %d does not support Store Slave Project CRC Parameter';
    16#30BB: F_EL6910MessageTemplate := 'if there are no Muting sensors behind the AOPD, the Backwards-Mode and optional Check of the OSSD inputs are not allowed';
    16#30BC: F_EL6910MessageTemplate := 'when optional Check of the OSSD inputs is activated, the Sequential Inputs mode has to be activated too';
    16#30BD: F_EL6910MessageTemplate := 'The number of Connections (%d) is unequal the calculated number of connections over all groups (%d)';
    16#30BE: F_EL6910MessageTemplate := 'The number of FBs (%d) is unequal the calculated number of FBs over all groups (%d)';
    16#30BF: F_EL6910MessageTemplate := 'The calculated local near process image size (%d) exceeded the maximum near local process image size of %d';
    16#30C0: F_EL6910MessageTemplate := 'the EtherCAT Output size was exceeded in the connection cfg data at word offset 0x%x (calculated value: %d, maximum value: %d)';
    16#30C1: F_EL6910MessageTemplate := 'the EtherCAT Input size was exceeded in the connection cfg data at word offset 0x%x (calculated value: %d, maximum value: %d)';
    16#30C2: F_EL6910MessageTemplate := 'the reserved bits in the flags of the Vendor Data were set (actual value: 0x%x, reserved flags: 0x%x)';
    16#30C3: F_EL6910MessageTemplate := 'FB CAMMON: if the Setting Mode is enabled, at least one position marker has to be configured in the cfg data';
    16#30C4: F_EL6910MessageTemplate := 'Connection Type is not supported at word-offset 0x%x of the cfg data';
    16#30C5: F_EL6910MessageTemplate := 'writing the PROFIsafe F-Parameter is not allowed in this logic state (%d), the logic state has to be 1 (RUN)';
    16#30C6: F_EL6910MessageTemplate := 'The ConnId 0x%x is used at least twice';
    16#30C7: F_EL6910MessageTemplate := 'The PROFIsafe Address 0x%x is used at least twice';
    16#30C8: F_EL6910MessageTemplate := 'The FSoE Address 0x%x is used at least twice';
    16#30C9: F_EL6910MessageTemplate := 'The TwinSAFE SC type %d is used at least twice';
    16#30CA: F_EL6910MessageTemplate := 'The TwinSAFE SC CRC 0x%x is used at least twice';
    16#30CB: F_EL6910MessageTemplate := 'The Connection Index %d in a FB Connection Shutdown is used at least twice';
    16#30CC: F_EL6910MessageTemplate := 'It is not allowed that the number of FBs and the number of Connections is zero inside the Group Cfg Data';
    16#30CD: F_EL6910MessageTemplate := 'the storing of the Store Slave Project CRC Parameter is not supported in connection %d';
    16#30CE: F_EL6910MessageTemplate := 'The received size of Safety Input Messages (%d) was too big, the maximum allowed value is %d';
    16#30CF: F_EL6910MessageTemplate := 'The received size of Safety Output Messages (%d) was too big, the maximum allowed value is %d';
    16#30D0: F_EL6910MessageTemplate := 'The received size of PROFIsafe Input Messages (%d) was too big, the maximum allowed value is %d';
    16#30D1: F_EL6910MessageTemplate := 'The received size of PROFIsafe Output Messages (%d) was too big, the maximum allowed value is %d';
    16#30D2: F_EL6910MessageTemplate := 'The Restore Mode is supported on a TwinSAFE SC connection at word-offset 0x%x';
    16#30D3: F_EL6910MessageTemplate := 'The FB %d (Connection Shutdown) is assigned to a non FSoE-connection';
    16#30D4: F_EL6910MessageTemplate := 'The download of the TwinSAFE IO-Project failed because %d FBs are configured (no FBs allowed)';
    16#30D5: F_EL6910MessageTemplate := 'When the TwinSAFE-Address in the Project Cfg data should be used, it has to be unequal zero';
    16#30D6: F_EL6910MessageTemplate := 'When the TwinSAFE-Address in the Project Cfg data should be used, the DIP-switch has to be zero (0x%x found)';
    16#30D7: F_EL6910MessageTemplate := 'Read aborted because of invalid code buffer offset (Calculated=0x%x, Expected=0x%x)';
    16#30D8: F_EL6910MessageTemplate := 'Invalid Safe User Parameter Offset at word offset 0x%x (Calculated=0x%x, Expected=0x%x)';
    16#30D9: F_EL6910MessageTemplate := 'The Standard Inputs Size of zero is not allowed';
    16#30DA: F_EL6910MessageTemplate := 'The download of the Replacement Values is not allowed after the download before (download state=%d)';
    16#30DB: F_EL6910MessageTemplate := 'The Info Data Map Cfg Data were downloaded in the wrong download state (%d)';
    16#30DC: F_EL6910MessageTemplate := 'The offset for the safety-Timer has to be inside the safety Output Area from 0x%x to 0x%x';
    16#30DD: F_EL6910MessageTemplate := 'The safety input size of connection %d is zero offset, the Safety Inputs cannot be mapped at byte offset 0x%x of Info Data Map Cfg Data';
    16#30DE: F_EL6910MessageTemplate := 'The safety output size of connection %d is zero, the Safety Outputs cannot be mapped at byte offset 0x%x of Info Data Map Cfg Data';
    16#30DF: F_EL6910MessageTemplate := 'No more safe user parameter expected at byte-offset 0x%x of the Safe User Parameter Cfg Data';
    16#30E0: F_EL6910MessageTemplate := 'The TwinSAFE Address 0 is not allowed in the Project Cfg Data';
    16#30E1: F_EL6910MessageTemplate := 'The download of the TwinSAFE IO-Project failed because %d Groups are configured (only 1 Group allowed)';
    16#30E2: F_EL6910MessageTemplate := 'The download of the Delete Project Cfg Data is not allowed in this state (%d)';
    16#30E3: F_EL6910MessageTemplate := 'The destination bit address (0x%x, Bit %d) already exists in the same mapping code';
    16#30E4: F_EL6910MessageTemplate := 'Local Inputs cannot be mapped in the Info data because no local inputs are existing';
    16#30E5: F_EL6910MessageTemplate := 'Local Outputs cannot be mapped in the Info data because no local outputs are existing';
    16#30E6: F_EL6910MessageTemplate := 'The destination bit address (0x%x, Bit %d) already exists in the same mapping code';
    16#30E7: F_EL6910MessageTemplate := 'the input mapping cfg data has to be read before the output mapping cfg data';
    16#30E8: F_EL6910MessageTemplate := 'wrong subindex order when reading the mapping cfg data, the expected subindex is %d';
    16#30E9: F_EL6910MessageTemplate := 'when reading the input mapping cfg data, it has to be started with subindex 1';
    16#30EA: F_EL6910MessageTemplate := 'invalid CRC when checking the Page %d of the Safe Logic Cfg Data';
    16#30EB: F_EL6910MessageTemplate := 'invalid CRC when checking the Page %d of the Safe User Parameter Cfg Data';
    16#30EC: F_EL6910MessageTemplate := 'invalid CRC when checking the Page %d of the Replacement values Cfg Data';
    16#3100: F_EL6910MessageTemplate := 'No groups defined when trying to activate or deactivate groups';
    16#3101: F_EL6910MessageTemplate := 'The reserved bits are set in value %d at offset %d when trying to activate or deactivate groups';
    16#3102: F_EL6910MessageTemplate := 'The operation mode at offset %d is not supported when trying to activate or deactivate groups';
    16#3103: F_EL6910MessageTemplate := 'The deactivation of groups is not enabled for any group so no replacement values should be downloaded';
    16#3104: F_EL6910MessageTemplate := 'The maximum number (%d) of Cfg Data pages was exceeded in the Replacement Values Cfg Data';
    16#3105: F_EL6910MessageTemplate := 'Invalid FB output size size at offset %d of the Replacement Values Cfg Data';
    16#3106: F_EL6910MessageTemplate := 'Unexpected groupindex in the Replacement values Cfg Data at offset 0x%x';
    16#3107: F_EL6910MessageTemplate := 'The download of the Activate Project Cfg Data was refused because %d bytes of the Replacement Values Cfg Data were missing';
    16#3108: F_EL6910MessageTemplate := 'To activate the Group %d the user has to logged in with access rights Bit 0-15 unequal 0 that the Safe Logic Program will be stopped when logging in';
    16#3109: F_EL6910MessageTemplate := 'No more definitions of individual replace values for analog FB Outputs in case of Group State unequal RUN are expected at offset %d';
    16#310A: F_EL6910MessageTemplate := 'The offset in the definitions of individual replace values for analog FB Outputs in case of Group State unequal RUN was wrong at offset %d';
    16#310B: F_EL6910MessageTemplate := 'The source process image offset of the Cyclic FRAM Data is outside the FB analog input area at offset %d';
    16#310C: F_EL6910MessageTemplate := 'The source process image offset of the Cyclic FRAM Data has to even at offset %d';
    16#310D: F_EL6910MessageTemplate := 'The size of the Cyclic FRAM Data was exceeding at offset %d';
    16#310E: F_EL6910MessageTemplate := 'The received size of the Cyclic FRAM Data at word offset 24 of the Safe Logic Cfg Data (%d) is unequal the calculated value of %d';
    16#310F: F_EL6910MessageTemplate := 'The size of the Cyclic FRAM CfgData in the GroupCfgData was not dividable by 4 at offset %d';
    16#3110: F_EL6910MessageTemplate := 'The offset of the Cyclic FRAM Data in the GroupCfgData was wrong at offset %d';
    16#3111: F_EL6910MessageTemplate := 'The value of %d at offset %d is not allowed when trying to activate or deactivate groups';
    16#3112: F_EL6910MessageTemplate := 'The activating or deactivating of groups is not allowed in PREOP';
    16#3113: F_EL6910MessageTemplate := 'FB CAMMON (Word-Offset 0x%x of the CfgData): The TDC2UpperLimit (%d) is lower or equal than the maximum position jitter (%d)';
    16#3114: F_EL6910MessageTemplate := 'FB CAMMON (Word-Offset 0x%x of the CfgData): The TDCUpperLimit (%d) is lower or equal than the maximum position jitter (%d)';
    16#3115: F_EL6910MessageTemplate := 'FB CAMMON (Word-Offset 0x%x of the CfgData): The value of TDCLowerLimit (plus maximum position jitter) (%d) is bigger or equal the configured position of 360 deg (%d)';
    16#3116: F_EL6910MessageTemplate := 'FB CAMMON (Word-Offset 0x%x of the CfgData): The value of BDCUpperLimit (plus twice the maximum position jitter) (%d) is bigger or equal the value of TDCLowerLimit (%d)';
    16#3117: F_EL6910MessageTemplate := 'FB CAMMON (Word-Offset 0x%x of the CfgData): The value of BDCUpperLimit (%d) is smaller or equal the configured value of 180 deg (plus maximum position jitter) (%d)';
    16#3118: F_EL6910MessageTemplate := 'FB CAMMON (Word-Offset 0x%x of the CfgData): The value of BDCLowerLimit (plus maximum position jitter) (%d) is greater or equal the configured value of 180 deg (%d)';
    16#3119: F_EL6910MessageTemplate := 'FB CAMMON (Word-Offset 0x%x of the CfgData): The value of OverrunMax (plus twice the maximum position jitter) (%d) is bigger or equal the value of BDCLowerLimit (%d)';
    16#311A: F_EL6910MessageTemplate := 'FB CAMMON (Word-Offset 0x%x of the CfgData): The value of TDCUpperLimit (plus twice the maximum position jitter) (%d) is bigger or equal the value of OverrunMax (%d)';
    16#311B: F_EL6910MessageTemplate := 'FB CAMMON (Word-Offset 0x%x of the CfgData): The value of TDC1UpperLimit (plus the maximum position jitter) (%d) is bigger or equal the configured position of 360 deg (%d)';
    16#311C: F_EL6910MessageTemplate := 'FB CAMMON (Word-Offset 0x%x of the CfgData): The value of TDC1LowerLimit (plus twice the maximum position jitter) (%d) is bigger or equal the value of TDC1UpperLimit (5d)';
    16#311D: F_EL6910MessageTemplate := 'FB CAMMON (Word-Offset 0x%x of the CfgData): The value of TDC2LowerLimit (plus twice the maximum position jitter) (%d) is bigger or equal the value of BDCLowerLimit (%d)';
    16#311E: F_EL6910MessageTemplate := 'FB CAMMON (Word-Offset 0x%x of the CfgData): The value of TDC2UpperLimit (plus twice the maximum position jitter) (%d) is bigger or equal the value of TDC2LowerLimit (%d)';
    16#311F: F_EL6910MessageTemplate := 'The maximum size of the Replacement Values was exceeded at Word-Offset 0x%x of the Group Cfg Data';
    16#3120: F_EL6910MessageTemplate := 'If no deactivation mode is enabled the offset of the replacement values shall be zero at Word-Offset 0x%x of the Group Cfg Data';
    16#3121: F_EL6910MessageTemplate := 'No more replacement values expected at byte-offset 0x%x of the Replacement Values Cfg Data';
    16#3122: F_EL6910MessageTemplate := 'The Download of the Project CRC is not allowed in PREOP';
    16#3201: F_EL6910MessageTemplate := 'The F_ParVersion in the F_Prm_Flag2 of the F-Parameter at Word-Offset 0x%x is unequal 1 (PROFIsafe V2)';
    16#3202: F_EL6910MessageTemplate := 'The F_CRC1 of the F-Parameter at Word-Offset 0x%x is wrong';
    16#3203: F_EL6910MessageTemplate := 'The F_CRC_Length in the F_Prm_Flag1 of the F-Parameter is wrong at Word-Offset 0x%x, the expected value is 0 (3 Bytes CRC2)';
    16#3206: F_EL6910MessageTemplate := 'The I-Parameter CRC in the F-Parameter is wrong at Word-Offset 0x%x';
    16#3207: F_EL6910MessageTemplate := 'The F_Block_ID in the F_Prm_Flag2 of the F-Parameter is wrong at Word-Offset 0x%x, the expected value is 0 (No F_iPar_CRC, no F_WD_Time 2) or 1 (F_iPar_CRC, no F_WD_Time 2)';
    16#3208: F_EL6910MessageTemplate := 'The F_Source_Address in the F-Parameter at Word-Offset 0x%x is outside the allowed area of 1-0xFFFE';
    16#3209: F_EL6910MessageTemplate := 'The F_Destination_Address in the F-Parameter at Word-Offset 0x%x is outside the allowed area of 1-0xFFFE';
    16#320A: F_EL6910MessageTemplate := 'The F_WD_Time in the F-parameter at Word-Offset 0x%x is outside the allowed range from 2-60000';
    16#320B: F_EL6910MessageTemplate := 'The F_Destination_Address in the F-Parameter at Word-Offset 0x%x is wrong, the expected value is %d';
    16#3300: F_EL6910MessageTemplate := 'The State OPERATIONAL was left in Restore Mode';
    16#3301: F_EL6910MessageTemplate := 'Only %d CRCs were matching in Restore Mode';
    16#3302: F_EL6910MessageTemplate := 'The CRC of the Activate Project Cfg Data in Restore Mode does not match, the expected value was 0x%x';
    16#3303: F_EL6910MessageTemplate := 'No RestoreMode Slaves configured when trying to start the Restore Mode';
    16#3304: F_EL6910MessageTemplate := 'The CRC of the User List Cfg Data was not matching in Restore Mode, the expected value was 0x%x';
    16#3305: F_EL6910MessageTemplate := 'The download of the User List Cfg Data is not activated in Restore Mode';
    16#3306: F_EL6910MessageTemplate := 'The download of the User List Cfg Data in Restore-Mode is not allowed in the state %d';
    16#3307: F_EL6910MessageTemplate := 'The activation of the TwinSAFE Restore Project is not allowed in the state %d';
    16#3308: F_EL6910MessageTemplate := 'The Restore Mode is not supported in EtherCAT state 0x%x';
    16#3310: F_EL6910MessageTemplate := 'The FSoE-Slave on the %d. connection is in Restore-Mode';
    16#3311: F_EL6910MessageTemplate := 'The FSoE-Master on the %d. connection is in Restore-Mode';
    16#3400: F_EL6910MessageTemplate := 'The %d. group has no more errors';
    16#3401: F_EL6910MessageTemplate := 'The Analog Input at word offset %d of the analog input process image has expired maximum allowed deviation to the last stored value, received value: %d, last stored value: %d';
    16#3402: F_EL6910MessageTemplate := 'The Wait-Com-Error-Timeout has not been expired when the group %d should be deactivated in passivate mode';
    16#3403: F_EL6910MessageTemplate := 'A module fault happened in group %d';
    16#3404: F_EL6910MessageTemplate := 'The assigned connection reported an error when the group %d was deactivated in passivate mode';
    16#3405: F_EL6910MessageTemplate := 'The connection has been successfully restarted when the group %d was deactivated in passivate mode';
    16#3410: F_EL6910MessageTemplate := 'All groups will enter the ERROR-state because the safe logic program has been restarted';
    16#3411: F_EL6910MessageTemplate := 'All groups will enter the ERROR-state because the CRC of the Change Group Activation Data was wrong';
    16#3412: F_EL6910MessageTemplate := 'All groups will enter the ERROR-state because the CRC of the Change FB Parameter Data was wrong';
    16#3413: F_EL6910MessageTemplate := 'All groups will enter the ERROR-state because the CRC of the Project CRC Data was wrong';
    16#3414: F_EL6910MessageTemplate := 'All groups will enter the ERROR-state because the CRC of the Cyclic FRAM Data was wrong';
    16#3415: F_EL6910MessageTemplate := 'The TwinSAFE Logic Program was not loaded on C1 because of an inconsistency';
    16#3416: F_EL6910MessageTemplate := 'The TwinSAFE Logic Program was not loaded on C2 because of an inconsistency';
    16#3417: F_EL6910MessageTemplate := 'All groups will enter the ERROR-state because the initialization of Cyclic FRAM Data was wrong';
    16#3418: F_EL6910MessageTemplate := 'Safe User Parameter from FRAM are not correct';
    16#3420: F_EL6910MessageTemplate := 'No more EtherCAT size error (EtherCAT Output Size=%d, EtherCAT Input Size=%d)';
    16#3421: F_EL6910MessageTemplate := 'The EtherCAT Output Data sizes of the Safety Logic Program (%d) and the EtherCAT Configuration (%d) are unequal';
    16#3422: F_EL6910MessageTemplate := 'The EtherCAT Input Data sizes of the Safety Logic Program (%d) and the EtherCAT Configuration (%d) are unequal';
    16#3423: F_EL6910MessageTemplate := 'The EtherCAT Output Data sizes for PROFIsafe of the Safety Logic Program (%d) and the EtherCAT Configuration (%d) are unequal';
    16#3424: F_EL6910MessageTemplate := 'The EtherCAT Input Data sizes for PROFIsafe of the Safety Logic Program (%d) and the EtherCAT Configuration (%d) are unequal';
    16#3425: F_EL6910MessageTemplate := 'The needed EtherCAT Process data buffer size (%d) exceeded the maximum available size of %d';
    16#3501: F_EL6910MessageTemplate := 'On the %d. connection the changeable FSoE Address of %d already exists';
    16#3502: F_EL6910MessageTemplate := 'On the %d. connection the changeable FSoE Address is zero';
    16#3800: F_EL6910MessageTemplate := 'FB %d (ESTOP): An EDM-fault (0x%x) was detected in state SAFE';
    16#3802: F_EL6910MessageTemplate := 'FB %d (ESTOP): An EDM-fault (0x%x) was detected in state RESET';
    16#3803: F_EL6910MessageTemplate := 'FB %d (ESTOP): An EDM-fault (0x%x) was detected in state START';
    16#3804: F_EL6910MessageTemplate := 'FB %d (ESTOP): An DiscTime-Fault (0x%x) was detected in state SAFE, the actual EStopIn-values are 0x%x';
    16#3806: F_EL6910MessageTemplate := 'FB %d (ESTOP): An DiscTime-Fault (0x%x) was detected in state RESET, the actual EStopIn-values are 0x%x';
    16#3807: F_EL6910MessageTemplate := 'FB %d (ESTOP): An DiscTime-Fault (0x%x) was detected in state START, the actual EStopIn-values are 0x%x';
    16#3809: F_EL6910MessageTemplate := 'FB %d (ESTOP): An DiscTime-Fault (0x%x) was detected in state DELAYOUT, the actual EStopIn-values are 0x%x';
    16#380F: F_EL6910MessageTemplate := 'FB %d (ESTOP): At least one activated EDM-Input was not reset in RUN when the EDM Reset time had been expired (Diag-Code=0x%x)';
    16#3810: F_EL6910MessageTemplate := 'FB %d (MON): An EDM-fault (0x%x) was detected in state SAFE';
    16#3812: F_EL6910MessageTemplate := 'FB %d (MON): An EDM-fault (0x%x) was detected in state RESET';
    16#3813: F_EL6910MessageTemplate := 'FB %d (MON): An EDM-fault (0x%x) was detected in state START';
    16#3814: F_EL6910MessageTemplate := 'FB %d (MON): An DiscTime-Fault (0x%x) was detected in state SAFE, the actual MonIn/Secure-values are 0x%x';
    16#3816: F_EL6910MessageTemplate := 'FB %d (MON): An DiscTime-Fault (0x%x) was detected in state RESET, the actual MonIn/Secure-values are 0x%x';
    16#3817: F_EL6910MessageTemplate := 'FB %d (MON): An DiscTime-Fault (0x%x) was detected in state START, the actual MonIn/Secure-values are 0x%x';
    16#3818: F_EL6910MessageTemplate := 'FB %d (MON): An DiscTime-Fault (0x%x) was detected in state RUN, the actual MonIn/Secure-values are 0x%x';
    16#3819: F_EL6910MessageTemplate := 'FB %d (MON): An DiscTime-Fault (0x%x) was detected in state DELAYOUT, the actual MonIn/Secure-values are 0x%x';
    16#381A: F_EL6910MessageTemplate := 'FB %d (MON): An DiscTime-Fault (0x%x) was detected in state FUNCTEST, the actual MonIn/Secure-values are 0x%x';
    16#381F: F_EL6910MessageTemplate := 'FB %d (MON): At least one activated EDM-Input was not reset in RUN when the EDM Reset time had been expired (Diag-Code=0x%x)';
    16#3820: F_EL6910MessageTemplate := 'FB %d (TWOHAND): A Disc-Group-fault (0x%x) was detected in state 1BUTTON, the actual TwoHandIn-values are 0x%x';
    16#3821: F_EL6910MessageTemplate := 'FB %d (TWOHAND): A Disc-Group-fault (0x%x) was detected in state 2BUTTON, the actual TwoHandIn-values are 0x%x';
    16#3823: F_EL6910MessageTemplate := 'FB %d (TWOHAND): An DiscTime-Fault (0x%x) was detected in state SAFE, the actual TwoHandIn-values are 0x%x';
    16#3825: F_EL6910MessageTemplate := 'FB %d (TWOHAND): An DiscTime-Fault (0x%x) was detected in state RESET, the actual TwoHandIn-values are 0x%x';
    16#382B: F_EL6910MessageTemplate := 'FB %d (TWOHAND): An DiscTime-Fault (0x%x) was detected in state 1BUTTON, the actual TwoHandIn-values are 0x%x';
    16#382C: F_EL6910MessageTemplate := 'FB %d (TWOHAND): An DiscTime-Fault (0x%x) was detected in state 2BUTTON, the actual TwoHandIn-values are 0x%x';
    16#382D: F_EL6910MessageTemplate := 'FB %d (TWOHAND): An DiscTime-Fault (0x%x) was detected in state RELEASE, the actual TwoHandIn-values are 0x%x';
    16#3830: F_EL6910MessageTemplate := 'FB %d (OPMODE): An DiscTime-Fault (0x%x) was detected, the actual OpIn-values are 0x%x';
    16#3831: F_EL6910MessageTemplate := 'FB %d (OPMODE): An Input-Fault was detected in state RESET, the actual OpIn-values are 0x%x';
    16#3840: F_EL6910MessageTemplate := 'FB %d (EDM): The SwitchOn-Time had been expired';
    16#3841: F_EL6910MessageTemplate := 'FB %d (EDM): The SwitchOff-Time had been expired';
    16#3853: F_EL6910MessageTemplate := 'FB %d (CS): An DiscTime-Fault (0x%x) was detected in state SAFE, the actual Deactivate-values are 0x%x';
    16#3855: F_EL6910MessageTemplate := 'FB %d (CS): An DiscTime-Fault (0x%x) was detected in state RESET, the actual Deactivate-values are 0x%x';
    16#3881: F_EL6910MessageTemplate := 'FB %d (MUTING): An DiscTime-Fault (0x%x) was detected in state RUN, the actual MuteIn/OssdIn-values are 0x%x';
    16#3883: F_EL6910MessageTemplate := 'FB %d (MUTING): An DiscTime-Fault (0x%x) was detected in state SAFE, the actual MuteIn/OssdIn-values are 0x%x';
    16#3885: F_EL6910MessageTemplate := 'FB %d (MUTING): An DiscTime-Fault (0x%x) was detected in state RESET, the actual MuteIn/OssdIn-values are 0x%x';
    16#3888: F_EL6910MessageTemplate := 'FB %d (MUTING): An DiscTime-Fault (0x%x) was detected in state DELAYOUT, the actual MuteIn/OssdIn-values are 0x%x';
    16#3889: F_EL6910MessageTemplate := 'FB %d (MUTING): An DiscTime-Fault (0x%x) was detected in state MUTING1, the actual MuteIn/OssdIn-values are 0x%x';
    16#388A: F_EL6910MessageTemplate := 'FB %d (MUTING): An DiscTime-Fault (0x%x) was detected in state MUTING2, the actual MuteIn/OssdIn-values are 0x%x';
    16#388B: F_EL6910MessageTemplate := 'FB %d (MUTING): An DiscTime-Fault (0x%x) was detected in state MUTING3, the actual MuteIn/OssdIn-values are 0x%x';
    16#388C: F_EL6910MessageTemplate := 'FB %d (MUTING): An DiscTime-Fault (0x%x) was detected in state MUTING4, the actual MuteIn/OssdIn-values are 0x%x';
    16#388D: F_EL6910MessageTemplate := 'FB %d (MUTING): An DiscTime-Fault (0x%x) was detected in state MUTING5, the actual MuteIn/OssdIn-values are 0x%x';
    16#388E: F_EL6910MessageTemplate := 'FB %d (MUTING): An DiscTime-Fault (0x%x) was detected in state MUTING6, the actual MuteIn/OssdIn-values are 0x%x';
    16#388F: F_EL6910MessageTemplate := 'FB %d (MUTING): An DiscTime-Fault (0x%x) was detected in state MUTING7, the actual MuteIn/OssdIn-values are 0x%x';
    16#3890: F_EL6910MessageTemplate := 'FB %d (MUTING): An DiscTime-Fault (0x%x) was detected in state MUTING8, the actual MuteIn/OssdIn-values are 0x%x';
    16#3891: F_EL6910MessageTemplate := 'FB %d (MUTING): An DiscTime-Fault (0x%x) was detected in state MUTING9, the actual MuteIn/OssdIn-values are 0x%x';
    16#3892: F_EL6910MessageTemplate := 'FB %d (MUTING): State RUN, Sequential Inputs=TRUE: MutingEnable is set and the MuteIn-signals are invalid, the actual MuteIn/OssdIn-values are 0x%x';
    16#3893: F_EL6910MessageTemplate := 'FB %d (MUTING): State RUN, Sequential Inputs=FALSE: MutingEnable is set and the MuteIn-signals are invalid, the actual MuteIn/OssdIn-values are 0x%x';
    16#3894: F_EL6910MessageTemplate := 'FB %d (MUTING): State MUTING1, MutingEnable is set and the OssdIn-signals are invalid, the actual MuteIn/OssdIn-values are 0x%x';
    16#3895: F_EL6910MessageTemplate := 'FB %d (MUTING): State MUTING1, MutingEnable is set and the MuteIn-signals are invalid, the actual MuteIn/OssdIn-values are 0x%x';
    16#3896: F_EL6910MessageTemplate := 'FB %d (MUTING): State MUTING2, MutingEnable is set and the MuteIn-signals before the AOPD are invalid, the actual MuteIn/OssdIn-values are 0x%x';
    16#3897: F_EL6910MessageTemplate := 'FB %d (MUTING): State MUTING2, MutingEnable is set and the MuteIn-signals after the AOPD are invalid, the actual MuteIn/OssdIn-values are 0x%x';
    16#3898: F_EL6910MessageTemplate := 'FB %d (MUTING): State MUTING3, MutingEnable is set and the OssdIn-signals are invalid, the actual MuteIn/OssdIn-values are 0x%x';
    16#3899: F_EL6910MessageTemplate := 'FB %d (MUTING): State MUTING3, Sequential Inputs=TRUE: MutingEnable is set and the MuteIn-signals are invalid, the actual MuteIn/OssdIn-values are 0x%x';
    16#389A: F_EL6910MessageTemplate := 'FB %d (MUTING): State MUTING3, Sequential Inputs=FALSE: MutingEnable is set and the MuteIn-signals are invalid, the actual MuteIn/OssdIn-values are 0x%x';
    16#389B: F_EL6910MessageTemplate := 'FB %d (MUTING): State MUTING4, MutingEnable is set and the OssdIn-signals are invalid, the actual MuteIn/OssdIn-values are 0x%x';
    16#389C: F_EL6910MessageTemplate := 'FB %d (MUTING): State MUTING4, MutingEnable is set and the MuteIn-signals are invalid, the actual MuteIn/OssdIn-values are 0x%x';
    16#389D: F_EL6910MessageTemplate := 'FB %d (MUTING): State MUTING5, MutingEnable is set and the OssdIn-signals are invalid, the actual MuteIn/OssdIn-values are 0x%x';
    16#389E: F_EL6910MessageTemplate := 'FB %d (MUTING): State MUTING5, Sequential Inputs=TRUE: MutingEnable is set and the MuteIn-signals are invalid, the actual MuteIn/OssdIn-values are 0x%x';
    16#389F: F_EL6910MessageTemplate := 'FB %d (MUTING): State MUTING5, Sequential Inputs=FALSE: MutingEnable is set and the MuteIn-signals are invalid, the actual MuteIn/OssdIn-values are 0x%x';
    16#38A0: F_EL6910MessageTemplate := 'FB %d (MUTING): State MUTING6, MutingEnable is set and the OssdIn-signals are invalid, the actual MuteIn/OssdIn-values are 0x%x';
    16#38A1: F_EL6910MessageTemplate := 'FB %d (MUTING): State MUTING6, MutingEnable is set and the MuteIn-signals are invalid, the actual MuteIn/OssdIn-values are 0x%x';
    16#38A2: F_EL6910MessageTemplate := 'FB %d (MUTING): State MUTING7, MutingEnable is set and the MuteIn-signals before the AOPD are invalid, the actual MuteIn/OssdIn-values are 0x%x';
    16#38A3: F_EL6910MessageTemplate := 'FB %d (MUTING): State MUTING7, MutingEnable is set and the MuteIn-signals after the AOPD are invalid, the actual MuteIn/OssdIn-values are 0x%x';
    16#38A4: F_EL6910MessageTemplate := 'FB %d (MUTING): State MUTING8, MutingEnable is set and the OssdIn-signals are invalid, the actual MuteIn/OssdIn-values are 0x%x';
    16#38A5: F_EL6910MessageTemplate := 'FB %d (MUTING): State MUTING8, Sequential Inputs=TRUE, CheckOssdOptional=TRUE: MutingEnable is set and the OssdIn-signals are invalid, the actual MuteIn/OssdIn-values are 0x%x';
    16#38A6: F_EL6910MessageTemplate := 'FB %d (MUTING): State MUTING8, Sequential Inputs=TRUE: MutingEnable is set and the MuteIn-signals are invalid, the actual MuteIn/OssdIn-values are 0x%x';
    16#38A7: F_EL6910MessageTemplate := 'FB %d (MUTING): State MUTING8, Sequential Inputs=FALSE: MutingEnable is set and the MuteIn-signals are invalid, the actual MuteIn/OssdIn-values are 0x%x';
    16#38A8: F_EL6910MessageTemplate := 'FB %d (MUTING): State MUTING9, MutingEnable is set and the OssdIn-signals are invalid, the actual MuteIn/OssdIn-values are 0x%x';
    16#38A9: F_EL6910MessageTemplate := 'FB %d (MUTING): State MUTING9, MutingEnable is set and the MuteIn-signals are invalid, the actual MuteIn/OssdIn-values are 0x%x';
    16#38AA: F_EL6910MessageTemplate := 'FB %d (MUTING): State MUTING5, Sequential Inputs=TRUE, MuteIn3 and MuteIn4 are inactive: MutingEnable is set and the MuteIn-signals are invalid, the actual MuteIn/OssdIn-values are 0x%x';
    16#38AB: F_EL6910MessageTemplate := 'FB %d (MUTING): State MUTING6, Sequential Inputs=TRUE, MuteIn3 and MuteIn4 are inactive: MutingEnable is set and the MuteIn-signals are invalid, the actual MuteIn/OssdIn-values are 0x%x';
    16#38AC: F_EL6910MessageTemplate := 'FB %d (MUTING): State MUTING1, MutingEnable is set and the MuteIn-signals are invalid, the actual MuteIn/OssdIn-values are 0x%x';
    16#38B0: F_EL6910MessageTemplate := 'FB %d (MUTING): At least one activated EDM-Input was not reset in RUN when the EDM Reset time had been expired (Diag-Code=0x%x)';
    16#38C1: F_EL6910MessageTemplate := 'FB %d (MUTING): The Max-Muting-Time had been expired in state MUTING1 (Digital Inputs=0x%x)';
    16#38C2: F_EL6910MessageTemplate := 'FB %d (MUTING): The Max-Muting-Time had been expired in state MUTING2 (Digital Inputs=0x%x)';
    16#38C3: F_EL6910MessageTemplate := 'FB %d (MUTING): The Max-Muting-Time had been expired in state MUTING3 (Digital Inputs=0x%x)';
    16#38C4: F_EL6910MessageTemplate := 'FB %d (MUTING): The Max-Muting-Time had been expired in state MUTING4 (Digital Inputs=0x%x)';
    16#38C5: F_EL6910MessageTemplate := 'FB %d (MUTING): The Max-Muting-Time had been expired in state MUTING5 (Digital Inputs=0x%x)';
    16#38C6: F_EL6910MessageTemplate := 'FB %d (MUTING): The Max-Muting-Time had been expired in state MUTING6 (Digital Inputs=0x%x)';
    16#38C7: F_EL6910MessageTemplate := 'FB %d (MUTING): The Max-Muting-Time had been expired in state MUTING7 (Digital Inputs=0x%x)';
    16#38C8: F_EL6910MessageTemplate := 'FB %d (MUTING): The Max-Muting-Time had been expired in state MUTING8 (Digital Inputs=0x%x)';
    16#38C9: F_EL6910MessageTemplate := 'FB %d (MUTING): The Max-Muting-Time had been expired in state MUTING9 (Digital Inputs=0x%x)';
    16#4001: F_EL6910MessageTemplate := 'FB %d (CAMMON): The TDC2UpperLimit (%d) is lower or equal than the maximum position jitter (%d)';
    16#4002: F_EL6910MessageTemplate := 'FB %d (CAMMON): The Position (%d) is bigger than the maximum position (plus the maximum position jitter) (%d)';
    16#4003: F_EL6910MessageTemplate := 'FB %d (CAMMON): The input OverrunCAM was FALSE in the top dead center area, the actual position is %d';
    16#4004: F_EL6910MessageTemplate := 'FB %d (CAMMON): The input OverrunCAM changed from FALSE to TRUE outside the area between BDCUpperLimit and TDCLowerLimit, the actual position is %d';
    16#4005: F_EL6910MessageTemplate := 'FB %d (CAMMON): The input OverrunCAM was TRUE in the area between OverrunMax and BDCUpperLimit, the actual position is %d';
    16#4006: F_EL6910MessageTemplate := 'FB %d (CAMMON): The input OverrunCAM changed from TRUE to FALSE outside the area between OverrunMax and BDCLowerLimit, the actual position is %d';
    16#4007: F_EL6910MessageTemplate := 'FB %d (CAMMON): The input UpwardsCAM was FALSE in the area between BDCUpperLimit and TDCLowerLimit, the actual position is %d';
    16#4008: F_EL6910MessageTemplate := 'FB %d (CAMMON): The input UpwardsCAM changed from FALSE to TRUE outside the area between BDCLowerLimit and TDCLowerLimit, the actual position is %d';
    16#4009: F_EL6910MessageTemplate := 'FB %d (CAMMON): The input UpwardsCAM changed from TRUE to FALSE outside the area between TDCLowerLimit and OverrunMax, the actual position is %d';
    16#400A: F_EL6910MessageTemplate := 'FB %d (CAMMON): The Position was moving while waiting for a rising edge of the input Reset in the state MOVE-STOP';
    16#400B: F_EL6910MessageTemplate := 'FB %d (CAMMON): The Position was moving while waiting for a falling edge of the input Reset in the state MOVE-START';
    16#400C: F_EL6910MessageTemplate := 'FB %d (CAMMON): The Position %d in the area between OverrunMax and BDCLowerLimit was detected in the state MOVE-UP';
    16#400D: F_EL6910MessageTemplate := 'FB %d (CAMMON): The Position has left the top dead center while waiting for a stop, the actual position is %d';
    16#400E: F_EL6910MessageTemplate := 'FB %d (CAMMON): The Position has been changed negative';
    16#400F: F_EL6910MessageTemplate := 'FB %d (CAMMON): The input UpwardsCAM was TRUE in the area between OverrunMax and BDCLowerLimit';
    16#4010: F_EL6910MessageTemplate := 'FB %d (CAMMON): The Position has a circle overflow in Pendulum Mode, actual position=%d, last position=%d';
    16#4011: F_EL6910MessageTemplate := 'FB %d (CAMMON): The Position has moved while waiting for a rising edge of the input Reset in Pendulum Mode, actual position=%d, compare position=%d';
    16#4012: F_EL6910MessageTemplate := 'FB %d (CAMMON): The Input BackwardsMove is TRUE while the Position is between 180 deg and 360 deg, the actual position is %d';
    16#4013: F_EL6910MessageTemplate := 'FB %d (CAMMON): The Input BackwardsMove is TRUE while the moving is clockwise';
    16#4014: F_EL6910MessageTemplate := 'FB %d (CAMMON): The Position has moved while waiting for a falling edge of the input Reset in Pendulum Mode, actual position=%d, last position=%d';
    16#4015: F_EL6910MessageTemplate := 'FB %d (CAMMON): The value of TDCLowerLimit (plus maximum position jitter) (%d) is bigger or equal the configured position of 360 deg (%d)';
    16#4016: F_EL6910MessageTemplate := 'FB %d (CAMMON): The value of BDCUpperLimit (plus twice the maximum position jitter) (%d) is bigger or equal the value of TDCLowerLimit (%d)';
    16#4017: F_EL6910MessageTemplate := 'FB %d (CAMMON): The value of BDCUpperLimit (%d) is smaller or equal the configured value of 180 deg (plus maximum position jitter) (%d)';
    16#4018: F_EL6910MessageTemplate := 'FB %d (CAMMON): The value of BDCLowerLimit (plus maximum position jitter) (%d) is greater or equal the configured value of 180 deg (%d)';
    16#4019: F_EL6910MessageTemplate := 'FB %d (CAMMON): The value of OverrunMax (plus twice the maximum position jitter) (%d) is bigger or equal the value of BDCLowerLimit (%d)';
    16#401A: F_EL6910MessageTemplate := 'FB %d (CAMMON): The value of TDCUpperLimit (plus twice the maximum position jitter) (%d) is bigger or equal the value of OverrunMax (%d)';
    16#401B: F_EL6910MessageTemplate := 'FB %d (CAMMON): The value of TDC1UpperLimit (plus the maximum position jitter) (%d) is bigger or equal the configured position of 360 deg (%d)';
    16#401C: F_EL6910MessageTemplate := 'FB %d (CAMMON): The value of TDC1LowerLimit (plus twice the maximum position jitter) (%d) is bigger or equal the value of TDC1UpperLimit (5d)';
    16#401D: F_EL6910MessageTemplate := 'FB %d (CAMMON): The value of TDC2LowerLimit (plus twice the maximum position jitter) (%d) is bigger or equal the value of BDCLowerLimit (%d)';
    16#401E: F_EL6910MessageTemplate := 'FB %d (CAMMON): The value of TDC2UpperLimit (plus twice the maximum position jitter) (%d) is bigger or equal the value of TDC2LowerLimit (%d)';
    16#401F: F_EL6910MessageTemplate := 'FB %d (CAMMON): The input PressStarted is TRUE and the position did not move after the PressStartedDelayTime';
    16#4020: F_EL6910MessageTemplate := 'FB %d (CAMMON): The input PressStarted is TRUE and the position has stopped after moving before';
    16#4021: F_EL6910MessageTemplate := 'FB %d (CAMMON): The input PressStarted is TRUE and the position has not moved enough, the actual position is %d, the compare position is %d';
    16#4022: F_EL6910MessageTemplate := 'FB %d (CAMMON), Pendulum Mode: The Position has changed contra clockwise while moving up clockwise (actual Position=%d, old Position=%d)';
    16#4023: F_EL6910MessageTemplate := 'FB %d (CAMMON), Pendulum Mode: The Position has changed clockwise while moving up contra clockwise (actual Position=%d, old Position=%d)';
    16#4024: F_EL6910MessageTemplate := 'FB %d (CAMMON): The Position was moving while waiting for a falling edge of the input Reset in the state WAIT-FOR_RESET';
    16#4025: F_EL6910MessageTemplate := 'FB %d (CAMMON): The TDCUpperLimit (%d) is lower or equal than the maximum position jitter (%d)';
    16#4080: F_EL6910MessageTemplate := 'FB %d (ADD/SUB): an underflow was detected, AnalogIn1=%d, AnalogIn2=%d';
    16#4081: F_EL6910MessageTemplate := 'FB %d (ADD/SUB): an overflow was detected, AnalogIn1=%d, AnalogIn2=%d';
    16#4088: F_EL6910MessageTemplate := 'FB %d (SPEED): an underflow was detected, actual Position=%d, old Position=%d';
    16#4089: F_EL6910MessageTemplate := 'FB %d (SPEED): an overflow was detected, actual Position=%d, old Position=%d';
    16#4090: F_EL6910MessageTemplate := 'FB %d (LIMIT): the minimum value (%d) is bigger than the maximum value (%d)';
    16#4098: F_EL6910MessageTemplate := 'FB %d (COMPARE): an underflow was detected on CompOut (%d), the minimum allowed value is %d';
    16#4099: F_EL6910MessageTemplate := 'FB %d (COMPARE): an overflow was detected on CompOut (%d), the maximum allowed value is %d';
    16#40A0: F_EL6910MessageTemplate := 'FB %d (MUL): an underflow was detected, AnalogIn1=%d, AnalogIn2=%d';
    16#40A1: F_EL6910MessageTemplate := 'FB %d (MUL): an overflow was detected, AnalogIn1=%d, AnalogIn2=%d';
    16#40A8: F_EL6910MessageTemplate := 'FB %d (DIV): an underflow was detected, AnalogIn1=%d, AnalogIn2=%d';
    16#40A9: F_EL6910MessageTemplate := 'FB %d (DIV): an overflow was detected, AnalogIn1=%d, AnalogIn2=%d';
    16#40B0: F_EL6910MessageTemplate := 'FB %d (SCALE): an underflow was detected, AnalogIn=%d';
    16#40B1: F_EL6910MessageTemplate := 'FB %d (SCALE): an overflow was detected, AnalogIn=%d';
    16#40B2: F_EL6910MessageTemplate := 'FB %d (SCALE): an overflow was detected after multiplication, AnalogIn=%d';
    16#40B3: F_EL6910MessageTemplate := 'FB %d (SCALE): an overflow was detected before division when rounding up the value, AnalogIn=%d';
    16#40B8: F_EL6910MessageTemplate := 'FB %d (COUNT): an underflow was detected on ActValue (%d)';
    16#40B9: F_EL6910MessageTemplate := 'FB %d (COUNT): an overflow was detected on ActValue (%d)';
    16#40C0: F_EL6910MessageTemplate := 'FB %d (SLI): an underflow was detected on ActValue (%d), the minimum allowed value is %d';
    16#40C1: F_EL6910MessageTemplate := 'FB %d (SLI): an overflow was detected on ActValue (%d), the maximum allowed value is %d';
    16#40C8: F_EL6910MessageTemplate := 'FB %d (ENVELOPE): an underflow was detected on InValue (%d), the minimum allowed value is %d';
    16#40C9: F_EL6910MessageTemplate := 'FB %d (ENVELOPE): an overflow was detected on InValue (%d), the maximum allowed value is %d';
    16#40CA: F_EL6910MessageTemplate := 'FB %d (ENVELOPE): an overflow error was detected on InValue (%d), InValue+Offset is bigger than the maximum allowed value';
    16#40CB: F_EL6910MessageTemplate := 'FB %d (ENVELOPE): the MaxTime was expired (InValue=%d)';
    16#40D0: F_EL6910MessageTemplate := 'FB %d (SLP): MultiturnPos_LL (%d) is bigger than MultiturnPos_UL (%d)';
    16#40D1: F_EL6910MessageTemplate := 'FB %d (SLP): MultiturnPos_LL=MultiturnPos_UL and SingleturnPos_LL (%d) is bigger than SingleturnPos_UL (%d)';
    16#40D8: F_EL6910MessageTemplate := 'FB %d (SBT): Brake-Test failed in state %d';
    16#40D9: F_EL6910MessageTemplate := 'FB %d (SBT): Brake-Test Interval expired in state %d';
    16#40DA: F_EL6910MessageTemplate := 'FB %d (SBT): Brake-Test failed, Actual Position Deviation=%d, Maximum Position Deviation=%dInterval expired in state %d';
ELSE F_EL6910MessageTemplate := CONCAT('Unknown EL6910 Text ID 0x', F_EL6910Hex(WORD_TO_ULINT(wTextId),4));
END_CASE

END_FUNCTION

(* stored: Version 1.1.0.1, ProductVersion 3.1.4026.18
   POU F_EL6910MessageTemplate: Id {db43890e-391e-4ef4-be3f-438f1c412a79}, SpecialFunc None *)
